(* IEC 61131-3 sources: SRCI_CLIENT_PLC/RobotLibrary/Library/Structures/AxesGroup/Parameter, 1 file *)

(* ---- AxesGroupParameter.st ---- *)
{attribute 'pack_mode' := '1'}
// -------------------------------------------------------------------------
//  SRCI Robot Library
// -------------------------------------------------------------------------
//
//  Object:      AxesGroupParameter
//  Author:      Thorsten Brach
//  Date:        2024-06-01
//
//  Description:
//
//
//  Copyright:
//    (C) 2024 Thorsten Brach. All rights reserved
//             Licensed under the MIT License.
//
//  Disclaimer:
//    This project is provided without any guarantee and can be used for
//    private and commercial purposes. Any use is at the user’s
//    own risk and responsibility.
//
// -------------------------------------------------------------------------
TYPE AxesGroupParameter :
STRUCT
  /// PLC specific data
  Plc            : AxesGroupParameterPlc;
  /// RC data read by the function "ReadRobotData" (see chapter 6.1.2)
  Rob            : AxesGroupParameterRob;

(*  /// Optional cyclic data configuration
  OptionalCyclic : AxesGroupParameterOptionalCyclic;
*)
END_STRUCT
END_TYPE
